// TIA Portal V20 export
TYPE "T_RCV_DATA"
   STRUCT
      TRCV : Struct
         IN : Struct
            READ : Bool;
            ID : CONN_OUC;
            LEN : UDInt;
            ADHOC : Bool;
            DATA : Array[0..254] of Char;
         END_STRUCT;
         OUT : Struct
            NDR : Bool;
            BYSY : Bool;
            ERROR : Bool;
            STATUS : Word;
            RCVD_LEN : DWord;
         END_STRUCT;
      END_STRUCT;
   END_STRUCT;
END_TYPE
